# EPICS substitutions: db/Beckhoff_7XXX/ecmcEX72XX_OPT_state.substitutions
file "ecmcEX72XX_OPT_state.template"
{
  pattern {CH_ID}
          {"$(OPT_CH_ID=01)"}
}
